Fanuc KAREL source: KD00071.KL

PROGRAM KD00071
%NOLOCKGROUP
VAR
  I: INTEGER
  J: INTEGER
  B: BOOLEAN
  R: REAL
  S: STRING[80]
BEGIN
  CONDITION[1]:
  WHEN DIN[1] = ON DO
    UNHOLD
  ENDCONDITION
END KD00071
